// TIA Portal V21 export
// export: Created 2026-11-10T07:35:06.8180898Z, ExportSetting WithDefaults, DisplayName Totally Integrated Automation Portal, DisplayVersion V21 Update 3, DisplayName STEP 7 Professional, DisplayVersion V21 Update 3, DisplayName STEP 7 Safety, DisplayVersion V21, DisplayName Tech WebApplication, DisplayVersion V21, DisplayName WinCC Basic/Comfort/Advanced, DisplayVersion V21 Update 3, DisplayName WinCC Unified, DisplayVersion V21 Update 3
FUNCTION_BLOCK "FB_Lad_ex056"   // FB20, LAD
{ S7_Optimized_Access := 'TRUE' }
VERSION : 0.1
// stored: AutoNumber true, IsIECCheckEnabled false, IsRetainMemResEnabled false, MemoryReserve 100, SetENOAutomatically false, UDAEnableTagReadback false
   VAR_INPUT
      v_req : Bool;
      v_mode : USInt;
      v_laddr : HW_DEVICE;
      v_ret_val : Int;
   END_VAR
   VAR_OUTPUT
      v_busy : Bool;
   END_VAR
BEGIN

REGION Network 1: D_ACT_DP - Activate/deactivate DP slaves
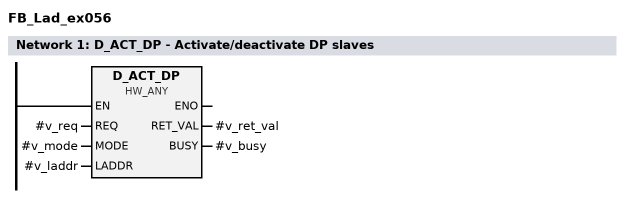
   RUNG wire#powerrail
      { S7_Templates := "[laddr_type := HW_ANY, mode_type := USInt]" } D_ACT_DP(REQ := #v_req, MODE := #v_mode, LADDR := #v_laddr, RET_VAL => #v_ret_val, BUSY => #v_busy)
   END_RUNG
   // the same network as SCL:
   #v_ret_val := D_ACT_DP(REQ := #v_req, MODE := #v_mode, LADDR := #v_laddr, BUSY => #v_busy);
END_REGION
END_FUNCTION_BLOCK
